RoboDK station: PickAndPlaceMultipart(Sriman).rdk

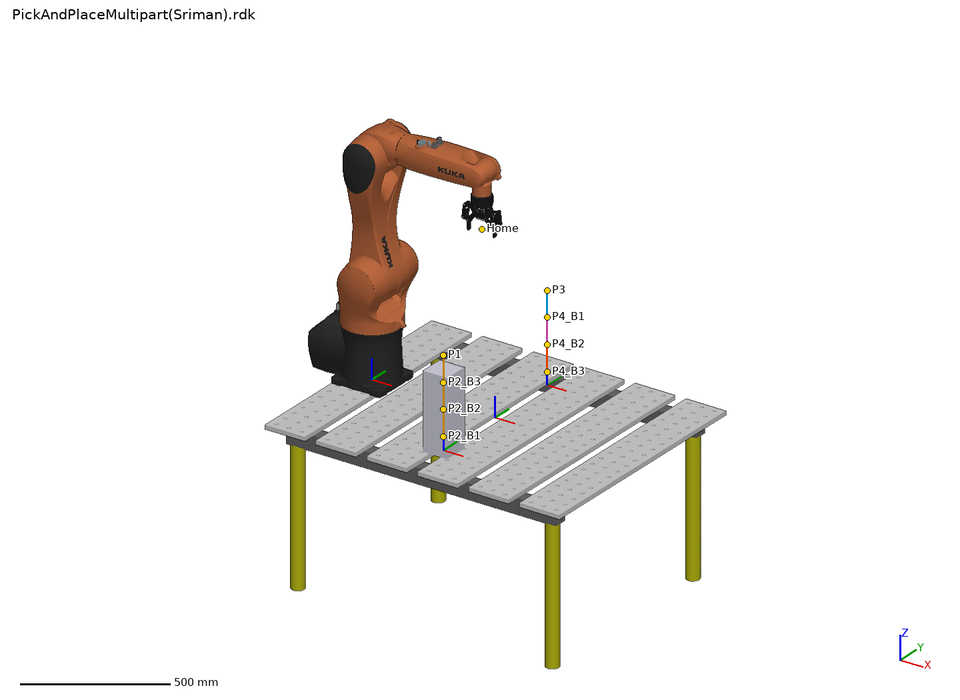
[picture v0: the station drawn from its stored meshes, robots at their saved joint values, targets as dots, program paths as lines]
Station PickAndPlaceMultipart(Sriman) (saved by RoboDK 6.1.1). Poses are relative to the parent item; angles as X-Y-Z fixed-axis rotations.
  - frame KUKA KR 10 R900 sixx Base at (0, 0, 0) mm
    - robot KUKA KR 10 R900 sixx: 6 axes, payload 10 kg, reach 901 mm, repeatability 0.03 mm, weight 52 kg
        modified DH rows (alpha deg, a mm, theta deg, d mm): 0, 0, 0, 400; -90, 25, 0, 0; 0, 455, -90, 0; -90, 35, 0, 420; 90, 0, 0, 0; -90, 0, 180, 80
        joint limits [-170, -190, -120, -185, -120, -350] to [170, 45, 156, 185, 120, 350]; home [0, -90, 90, 0, 0, 0]; saved at [0, -90, 90, 0, 90, 0]
      - tool RobotiQ 2F-85 Gripper (Open), TCP at (0, 0, 130) mm, size 147.4 x 75 x 146.8 mm
  - frame Base at (500, 0, 0) mm
    - object Table 1200x1000mm (Welding) at (0, 0, 0) mm, size 1193.8 x 965.2 x 609.6 mm, geometry from Table-1200x1000mm-Welding.sld
    - target Home (Cartesian target) at (-55, 0, 680) mm, rotated rx 180 ry 0 rz -180 deg; joints [0, -90, 90, 0, 90, 0] of KUKA KR 10 R900 sixx
  - frame Part1 at (500, -300, 0) mm
    - target P2_B3 (Cartesian target) at (0, 0, 250) mm, rotated rx 180 ry 0 rz 180 deg; joints [30.964, -53.73, 105.216, 0, 38.514, 30.964] of KUKA KR 10 R900 sixx
    - target P1 (Cartesian target) at (0, 0, 350) mm, rotated rx 180 ry 0 rz 180 deg; joints [30.964, -62.078, 101.89, 0, 50.188, 30.964] of KUKA KR 10 R900 sixx
    - target P2_B2 (Cartesian target) at (0, 0, 150) mm, rotated rx 180 ry 0 rz -180 deg; joints [30.964, -43.632, 105.52, 0, 28.112, 30.964] of KUKA KR 10 R900 sixx
    - target P2_B1 (Cartesian target) at (0, 0, 50) mm, rotated rx 180 ry 0 rz -180 deg; joints [30.964, -32.411, 102.794, 0, 19.616, 30.964] of KUKA KR 10 R900 sixx
    - object box1 at (0, 0, 50) mm, size 100 x 100 x 100 mm, geometry from box.sld
    - object box2 at (0, 0, 150) mm, size 100 x 100 x 100 mm, geometry from box.sld
    - object box3 at (0, 0, 250) mm, size 100 x 100 x 100 mm, geometry from box.sld
  - frame Part2 at (500, 300, 0) mm
    - target P3 (Cartesian target) at (0, 0, 350) mm, rotated rx 180 ry 0 rz -180 deg; joints [-30.964, -62.078, 101.89, 0, 50.188, -30.964] of KUKA KR 10 R900 sixx
    - target P4_B3 (Cartesian target) at (0, 0, 50) mm, rotated rx 180 ry 0 rz 180 deg; joints [-30.964, -32.411, 102.794, 0, 19.616, -30.964] of KUKA KR 10 R900 sixx
    - target P4_B2 (Cartesian target) at (0, 0, 150) mm, rotated rx 180 ry 0 rz 180 deg; joints [-30.964, -43.632, 105.52, 0, 28.112, -30.964] of KUKA KR 10 R900 sixx
    - target P4_B1 (Cartesian target) at (0, 0, 250) mm, rotated rx 180 ry 0 rz -180 deg; joints [-30.964, -53.73, 105.216, 0, 38.514, -30.964] of KUKA KR 10 R900 sixx
  - program Restore (1 instructions, listed below)
  - program Pick of box 3 (6 instructions, listed below)
  - program Place of Box 3 (6 instructions, listed below)
  - program Pick of box2 (6 instructions, listed below)
  - program Place of box 2 (6 instructions, listed below)
  - program Pick of box 1 (6 instructions, listed below)
  - program Place of box 1 (6 instructions, listed below)
  - program Main (7 instructions, listed below)
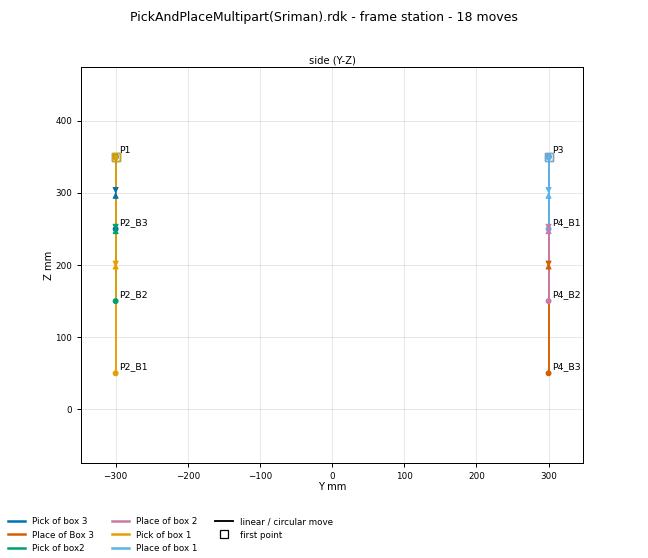
[picture p0: tool path of PickAndPlaceMultipart(Sriman).rdk in frame station, 18 of 18 moves have a stored position in this frame; points joined in program order, loops and branches not executed]

--- program Restore (robot KUKA KR 10 R900 sixx) ---
  Move objects

--- program Pick of box 3 (robot KUKA KR 10 R900 sixx) ---
  Set Ref.: Part1
  Set Tool: RobotiQ 2F-85 Gripper (Open)
  MoveJ (P1)
  MoveL (P2_B3)
  Attach to RobotiQ 2F-85 Gripper (Open)
  MoveL (P1)

--- program Place of Box 3 (robot KUKA KR 10 R900 sixx) ---
  Set Ref.: Part2
  Set Tool: RobotiQ 2F-85 Gripper (Open)
  MoveJ (P3)
  MoveL (P4_B3)
  Detach from RobotiQ 2F-85 Gripper (Open)
  MoveL (P3)

--- program Pick of box2 (robot KUKA KR 10 R900 sixx) ---
  Set Ref.: Part1
  Set Tool: RobotiQ 2F-85 Gripper (Open)
  MoveJ (P1)
  MoveL (P2_B2)
  Attach to RobotiQ 2F-85 Gripper (Open)
  MoveL (P1)

--- program Place of box 2 (robot KUKA KR 10 R900 sixx) ---
  Set Ref.: Part2
  Set Tool: RobotiQ 2F-85 Gripper (Open)
  MoveJ (P3)
  MoveL (P4_B2)
  Detach from RobotiQ 2F-85 Gripper (Open)
  MoveL (P3)

--- program Pick of box 1 (robot KUKA KR 10 R900 sixx) ---
  Set Ref.: Part1
  Set Tool: RobotiQ 2F-85 Gripper (Open)
  MoveJ (P1)
  MoveL (P2_B1)
  Attach to RobotiQ 2F-85 Gripper (Open)
  MoveL (P1)

--- program Place of box 1 (robot KUKA KR 10 R900 sixx) ---
  Set Ref.: Part2
  Set Tool: RobotiQ 2F-85 Gripper (Open)
  MoveJ (P3)
  MoveL (P4_B1)
  Detach from RobotiQ 2F-85 Gripper (Open)
  MoveL (P3)

--- program Main (robot KUKA KR 10 R900 sixx) ---
  Call Pick of box 3
  Call Place of Box 3
  Call Pick of box2
  Call Place of box 2
  Call Pick of box 1
  Call Place of box 1
  Call Restore
